Yaskawa INFORM job: HOME_TRACK.JBI

/JOB
//NAME HOME_TRACK
//POS
///NPOS 2,2,2,0,0,0
///TOOL 0
///POSTYPE PULSE
///PULSE
C00000=-283,-101162,-84213,3710,-80188,-1936
C00001=-283,-101162,-84213,3710,-80188,-1936
BC00000=570125
BC00001=570125
EC00000=192,0
EC00001=-2638,-94527
//INST
///DATE 2026/09/15 00:00
///ATTR SC,RW
///GROUP1 RB1,BS1
///GROUP2 ST1
NOP
MOVJ C00000 BC00000 VJ=20.00 DEC=20  +MOVJ EC00000 VJ=20.00
MOVJ C00001 BC00001 VJ=20.00 DEC=20  +MOVJ EC00001 VJ=20.00
END
